(* CODESYS project Elevator_Control.project

Project tree, tasks and I/O mapping:
  Device : CODESYS Control Win V3, CODESYS, version 3.5.21.0
    application Application
      libraries: Standard, 3.5.18.0 (System)
      task MainTask (cyclic, interval 70 ms, priority 1) calls PLC_PRG, Simulation, GA_Collector
      task VISU_TASK (cyclic, interval 100 ms, priority 31) calls VisuElems.Visu_Prg
      global variables GVL
      visualisation Visualization
      program Simulation [ST]
      program GA_Collector [FBD]
      program PLC_PRG [SFC]: _aOpeningDoor_exit, _aCallsHMI_active, _aClosingDoor_active_1, _aClosingDoor_exit_1, _aOpeningDoor_active_1, _aOpenDoor_active, _aClosingDoor_exit_1_1_1_1_1, _aHoming_exit, _aHoming_active, _aOpeningDoor_active_1_1, _aOpeningDoor_exit_1, _aClosingDoor1_exit, _aClosingDoor1_active, _aClosingDoor_active_1_1_1_1_1, _aOpenDoor_exit, _aOpenDoor1_active, _aOpenDoor1_exit, _aTargetMoveStart_active, _aTargetMoveStart_exit, _aOpenDoor2_active, _aOpenDoor2_exit, _aResetCalls_active
      ENUMs/
        GAs/
          data type State_GA
          data type Action_State
          data type DoWhats_Closing
          data type DoWhats_Opening
          data type DoWhats_Motor
        data type Fault
        data type SensorSequence
      GAs/
        function block Opening_GA [SFC]: _aInit_active, _aReady_active, _aBusy_active, _aOpeningDoor_active, _aEnd_active, _aEnd_exit, _aOpeningDoor_exit
        function block Closing_GA [SFC]: _aInit_active, _aCheckPresence_active, _aBusy_active, _aClosingDoor_active, _aClosingDoor_exit, _aEnd_active, _aEnd_exit, _aReady_active_1
        function block Motor_GA [SFC]: _aBusy_active, _aEnd_Cycle_active, _aEnd_INIT_exit, _aInit_active, _aReady_active, _aEnd_Cycle_exit, _aMotor_ON_active, _aSetting_Down_active, _aMovingElevator_active, _aSetting_Init_active, _aSetting_Up_active, _aUpdateFloor_active_1, _aEnd_INIT_active, _aChangeDirection_exit, _aChangeDirection_active, _aMovingElevator_exit, _aSequenceCheck_active, _aMoveFast_entry_1, _aUpdateFloor_entry_1, _aInvertedSpeed1_active, _aInvertedSpeed_active_1, _aInvertedSpeed_exit, _aInvertedSpeed_entry
  text list GlobalTextList
*)

// Device/Application/ENUMs/GAs/State_GA
//{attribute 'qualified_only'}
//{attribute 'strict'}
TYPE State_GA :
(
	S_Init,
	S_Ready,
	S_Busy
);
END_TYPE

// Device/Application/ENUMs/GAs/Action_State
//{attribute 'qualified_only'}
//{attribute 'strict'}
TYPE Action_State :
(
	Do_Action,
	WaitDone,
	SetOpOk
);
END_TYPE

// Device/Application/ENUMs/Fault
//{attribute 'qualified_only'}
//{attribute 'strict'}
TYPE Fault :
(
	None,
	MagnetRamp,
	MagnetDeck
);
END_TYPE

// Device/Application/ENUMs/SensorSequence
//{attribute 'qualified_only'}
//{attribute 'strict'}
TYPE SensorSequence :
(
	Seq_Deck,
	Seq_Ramp1,
	Seq_Ramp2,
	Seq_Fault
);
END_TYPE

// Device/Application/ENUMs/GAs/DoWhats_Closing
//{attribute 'qualified_only'}
//{attribute 'strict'}
TYPE DoWhats_Closing :
(
	Do_CloseDoor
);
END_TYPE

// Device/Application/ENUMs/GAs/DoWhats_Opening
//{attribute 'qualified_only'}
//{attribute 'strict'}
TYPE DoWhats_Opening :
(
	Do_OpenDoor
);
END_TYPE

// Device/Application/ENUMs/GAs/DoWhats_Motor
//{attribute 'qualified_only'}
//{attribute 'strict'}
TYPE DoWhats_Motor :
(
	Do_Up,
	Do_Down, 
	Do_Inizialization
);
END_TYPE

// Device/Application/GVL
//{attribute 'qualified_only'}
VAR_GLOBAL
(* Elevator managing variables*)
	Open: BOOL;				(* Sensor: the door is fully open*)
	Closed: BOOL;			(* Sensor: the door is fully closed*)
	LimitDown: BOOL;		(* Sensor: lower limit sensor, if TRUE the lift has reached the lower limit*)
	LimitUp: BOOL;			(* Sensor: upper limit sensor, if TRUE the lift has reached the upper limit*)
	DeckSensor: BOOL;		(* Sensor: if TRUE the cab is in proximity of a deck*)
	RampSensor: BOOL;		(* Sensor: if TRUE the cab is in proximity of a ramp*)
	Presence :BOOL; 		(* Sensor: if TRUE something blocks the door photocell*)
	Emergency: BOOL;		(* Input: if TRUE the emergency button has been pressed*)

	Closing: BOOL;			(* Actuator: if TRUE the door starts closing*)
	Opening: BOOL;			(* Actuator: the door starts opening*)
	Motor_on: BOOL;			(* Actuator: if TRUE the lift pulley motor start moving*)
	Up: BOOL;				(* Actuator parameter: if TRUE the lift moves upward, downward otherwise*)
	Vel: BOOL;				(* Actuator parameter: motor speed, if TRUE high speed, low speed otherwise*)


	Current: INT;  			(* Visualization: variable used to storage the current deck*)
    Destination: INT;		(* Visualization: variable used to storage the the destination deck*)
	EmergencyVis: BOOL; 	(* Visualization: if TRUE the emergency light is turned on*)

	InitialDeck: INT := 1;	(* Only for simulation: variable used to define the initial deck*)
	InitCycle: BOOL := FALSE;(* Only for simulation: used to execute the instruction at the first cycle*)
	Height: INT;			(* Only for simulation: elevator height*)
	DeckRest: INT;        	(* Only for simulation: division rest for generating deck sensor*)
	Memory: INT;
	RampRest: INT;			(* Only for simulation: division rest for generating the ramp position*)
	MemoryR: INT;
	Door: INT;				(* Only for simulation: to visualize the closing of the door*)
	Displacement: INT;		(* Only for simulation: lift displacement, dependent on the motor speed*)

 (*Inputs: internal panel variables*)
	PG: BOOL;
	P1: BOOL;
	P2: BOOL;
	P3: BOOL;
	P4: BOOL;
	P5: BOOL;
	P6: BOOL;
	P7: BOOL;

(*Visualization: internal panel variables used to turn on the LED*)
	PGVis: BOOL;
	P1Vis: BOOL;
	P2Vis: BOOL;
	P3Vis: BOOL;
	P4Vis: BOOL;
	P5Vis: BOOL;
	P6Vis: BOOL;
	P7Vis: BOOL;

(*Inputs: external panel variables*)
	UpDeckG: BOOL;
	UpDeck1: BOOL;
	UpDeck2: BOOL;
	UpDeck3: BOOL;
	UpDeck4: BOOL;
	UpDeck5: BOOL;
	UpDeck6: BOOL;
	DownDeck7: BOOL;
	DownDeck6: BOOL;
	DownDeck5: BOOL;
	DownDeck4: BOOL;
	DownDeck3: BOOL;
	DownDeck2: BOOL;
	DownDeck1: BOOL;

(*Visualization: external panel variables used to turn on the LED*)
	UpDeckGVis: BOOL;
	UpDeck1Vis: BOOL;
	UpDeck2Vis: BOOL;
	UpDeck3Vis: BOOL;
	UpDeck4Vis: BOOL;
	UpDeck5Vis: BOOL;
	UpDeck6Vis: BOOL;
	DownDeck7Vis: BOOL;
	DownDeck6Vis: BOOL;
	DownDeck5Vis: BOOL;
	DownDeck4Vis: BOOL;
	DownDeck3Vis: BOOL;
	DownDeck2Vis: BOOL;
	DownDeck1Vis: BOOL;

(*Only for simulation: variables used to simulate the fault on deck sensor*)
	SensorG: BOOL;				(* if TRUE the magnetic information for deck G is lost and the deck sensor cannot become TRUE*)
	Sensor1: BOOL;				(* if TRUE the magnetic information for deck 1 is lost and the deck sensor cannot become TRUE*)
	Sensor2: BOOL;
	Sensor3: BOOL;
	Sensor4: BOOL;
	Sensor5: BOOL;
	Sensor6: BOOL;
	Sensor7: BOOL;
	FaultSensorAlarm: BOOL; 	(* Visulaization: if TRUE alerts the user of a deck sensor fault*)

(*Only for simulation: variables used to simulate the fault on ramp sensor*)
	RampGUp: BOOL;
	Ramp1Down: BOOL;
	Ramp1Up:BOOL;
	Ramp2Down: BOOL;
	Ramp2Up:BOOL;
	Ramp3Down: BOOL;
	Ramp3Up:BOOL;
	Ramp4Down: BOOL;
	Ramp4Up:BOOL;
	Ramp5Down: BOOL;
	Ramp5Up:BOOL;
	Ramp6Down: BOOL;
	Ramp6Up:BOOL;
	Ramp7Down: BOOL;
	FaultRampAlarm: BOOL; 		(* Visulaization: if TRUE alerts the user of a ramp sensor fault*)
	SensorGOK: BOOL;
	Sensor1OK: BOOL;
	Sensor2OK: BOOL;
	Sensor6OK: BOOL;
	Sensor3OK: BOOL;
	Sensor4OK: BOOL;
	Sensor5OK: BOOL;
	Sensor7OK: BOOL;
	RampGUpOK: BOOL;
	Ramp1DownOK: BOOL;
	Ramp1UpOK: BOOL;
	Ramp2DownOK: BOOL;
	Ramp2UpOK: BOOL;
	Ramp3DownOK: BOOL;
	Ramp3UpOK: BOOL;
	Ramp4DownOK: BOOL;
	Ramp4UpOK: BOOL;
	Ramp5DownOK: BOOL;
	Ramp5UpOK: BOOL;
	Ramp6DownOK: BOOL;
	Ramp6UpOK: BOOL;
	Ramp7DownOK: BOOL;
	Ramp7UpOK: BOOL;
	
	Closing_GA_0: Closing_GA;
	Opening_GA_0: Opening_GA;
	Motor_GA_0: Motor_GA;
END_VAR

// Device/Application/PLC_PRG
PROGRAM PLC_PRG
VAR
	A_State: Action_State := Do_Action;
	OpOk: BOOL;
	IntPanel : ARRAY [0..7] OF BOOL;
	ExtPanelUP : ARRAY [0..6] OF BOOL;
	ExtPanelDOWN : ARRAY [1..7] OF BOOL;
	CallInt : ARRAY[0..7] OF BOOL; //chiamate interne
	CallUp : ARRAY[0..6] OF BOOL;     //chiamate esterne vs alto
	CallDown : ARRAY[1..7] OF BOOL;   //chiamate esterne vs basso   
	i : INT;
END_VAR

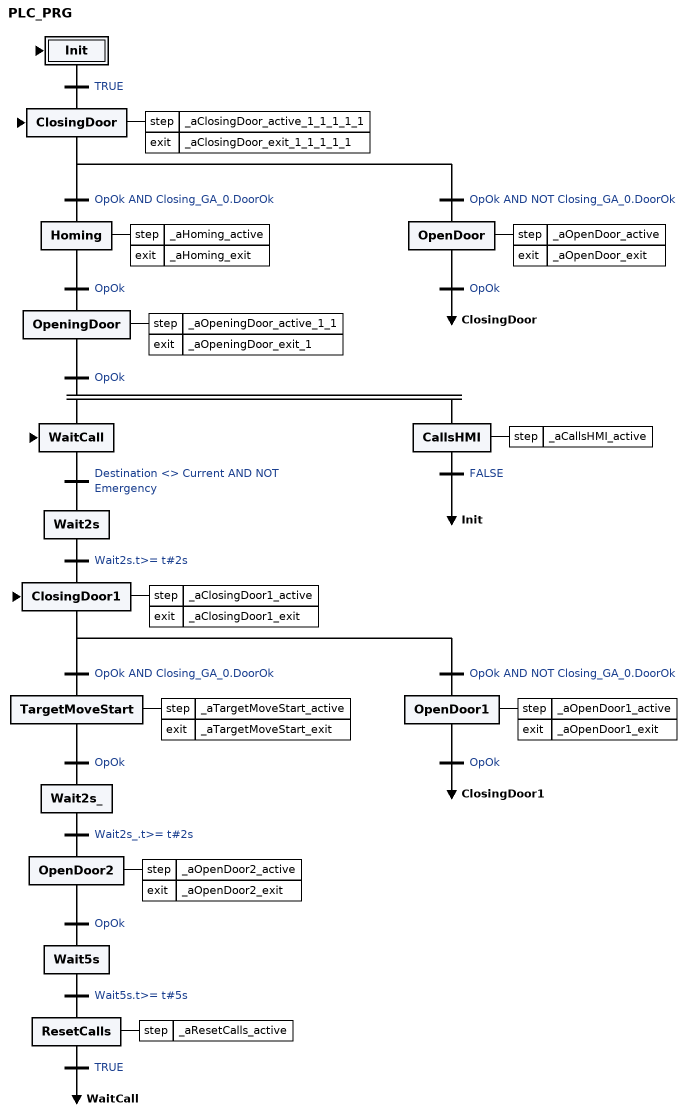
INITIAL_STEP Init:
END_STEP
TRANSITION FROM Init TO ClosingDoor
    := TRUE;
END_TRANSITION
STEP ClosingDoor:
    _aClosingDoor_active_1_1_1_1_1(N);  // step action
    _aClosingDoor_exit_1_1_1_1_1(P0);  // exit action
END_STEP
TRANSITION FROM ClosingDoor TO Homing
    := OpOk AND Closing_GA_0.DoorOk;
END_TRANSITION
TRANSITION FROM ClosingDoor TO OpenDoor
    := OpOk AND NOT Closing_GA_0.DoorOk;
END_TRANSITION
STEP OpenDoor:
    _aOpenDoor_active(N);  // step action
    _aOpenDoor_exit(P0);  // exit action
END_STEP
TRANSITION FROM OpenDoor TO ClosingDoor
    := OpOk;
END_TRANSITION
STEP Homing:
    _aHoming_active(N);  // step action
    _aHoming_exit(P0);  // exit action
END_STEP
TRANSITION FROM Homing TO OpeningDoor
    := OpOk;
END_TRANSITION
STEP OpeningDoor:
    _aOpeningDoor_active_1_1(N);  // step action
    _aOpeningDoor_exit_1(P0);  // exit action
END_STEP
TRANSITION FROM OpeningDoor TO (WaitCall, CallsHMI)
    := OpOk;
END_TRANSITION
STEP WaitCall:
END_STEP
STEP CallsHMI:
    _aCallsHMI_active(N);  // step action
END_STEP
TRANSITION FROM CallsHMI TO Init
    := FALSE;
END_TRANSITION
TRANSITION FROM WaitCall TO Wait2s
    := Destination <> Current AND NOT Emergency;
END_TRANSITION
STEP Wait2s:
END_STEP
TRANSITION FROM Wait2s TO ClosingDoor1
    := Wait2s.t>= t#2s;
END_TRANSITION
STEP ClosingDoor1:
    _aClosingDoor1_active(N);  // step action
    _aClosingDoor1_exit(P0);  // exit action
END_STEP
TRANSITION FROM ClosingDoor1 TO TargetMoveStart
    := OpOk AND Closing_GA_0.DoorOk;
END_TRANSITION
TRANSITION FROM ClosingDoor1 TO OpenDoor1
    := OpOk AND NOT Closing_GA_0.DoorOk;
END_TRANSITION
STEP OpenDoor1:
    _aOpenDoor1_active(N);  // step action
    _aOpenDoor1_exit(P0);  // exit action
END_STEP
TRANSITION FROM OpenDoor1 TO ClosingDoor1
    := OpOk;
END_TRANSITION
STEP TargetMoveStart:
    _aTargetMoveStart_active(N);  // step action
    _aTargetMoveStart_exit(P0);  // exit action
END_STEP
TRANSITION FROM TargetMoveStart TO Wait2s_
    := OpOk;
END_TRANSITION
STEP Wait2s_:
END_STEP
TRANSITION FROM Wait2s_ TO OpenDoor2
    := Wait2s_.t>= t#2s;
END_TRANSITION
STEP OpenDoor2:
    _aOpenDoor2_active(N);  // step action
    _aOpenDoor2_exit(P0);  // exit action
END_STEP
TRANSITION FROM OpenDoor2 TO Wait5s
    := OpOk;
END_TRANSITION
STEP Wait5s:
END_STEP
TRANSITION FROM Wait5s TO ResetCalls
    := Wait5s.t>= t#5s;
END_TRANSITION
STEP ResetCalls:
    _aResetCalls_active(N);  // step action
END_STEP
TRANSITION FROM ResetCalls TO WaitCall
    := TRUE;
END_TRANSITION

ACTION _aOpeningDoor_exit:
OpOk := FALSE;
A_State := Do_Action;
END_ACTION

ACTION _aCallsHMI_active:
// Mappatura dei tasti della pulsantiera interna sui piani
IntPanel[0] := PG;
IntPanel[1] := P1;
IntPanel[2] := P2;
IntPanel[3] := P3;
IntPanel[4] := P4;
IntPanel[5] := P5;
IntPanel[6] := P6;
IntPanel[7] := P7;

//Gestione delle richieste interne
FOR i := 0 TO 7 DO
	IF IntPanel[i] THEN
		CallInt[i] := TRUE;   	//Salva richiesta interna attiva
	END_IF
	IF (Current = i) AND Open THEN
		CallInt[i] := FALSE;   // Cancella richiesta se cabina è ferma al piano e porte aperte
	END_IF
END_FOR

// Mappatura dei tasti di salita della pulsantiera esterna
ExtPanelUP[0] := UpDeckG;
ExtPanelUP[1] := UpDeck1;
ExtPanelUP[2] := UpDeck2;
ExtPanelUP[3] := UpDeck3;
ExtPanelUP[4] := UpDeck4;
ExtPanelUP[5] := UpDeck5;
ExtPanelUP[6] := UpDeck6;

//Gestione delle richieste esterne verso l'alto
FOR i:= 0 TO 6 DO
	IF ExtPanelUP[i] THEN 
		CallUp[i] := TRUE;        
	END_IF;
	IF (Current = i) AND Open THEN
	CallUp[i] := FALSE;           
	END_IF
END_FOR

// Mappatura dei tasti di discesa della pulsantiera esterna
ExtPanelDOWN[1] := DownDeck1;
ExtPanelDOWN[2] := DownDeck2;
ExtPanelDOWN[3] := DownDeck3;
ExtPanelDOWN[4] := DownDeck4;
ExtPanelDOWN[5] := DownDeck5;
ExtPanelDOWN[6] := DownDeck6;
ExtPanelDOWN[7] := DownDeck7;

// Gestione delle richieste esterne verso il basso
FOR i := 1 TO 7 DO
	IF ExtPanelDown[i] THEN
		CallDown[i] := TRUE;
	END_IF
	IF (Current = i) AND Open THEN
	CallDown[i] := FALSE;
	END_IF
END_FOR

//Aggiornamento LED interni in base alle richieste
PGVis := CallInt[0];
P1Vis := CallInt[1];
P2Vis := CallInt[2];
P3Vis := CallInt[3];
P4Vis := CallInt[4];
P5Vis := CallInt[5];
P6Vis := CallInt[6];
P7Vis := CallInt[7];

//Aggiornamento LED esterni salita
UpDeckGVis := CallUp[0];
UpDeck1Vis := CallUp[1];
UpDeck2Vis := CallUp[2];
UpDeck3Vis := CallUp[3];
UpDeck4Vis := CallUp[4];
UpDeck5Vis := CallUp[5];
UpDeck6Vis := CallUp[6];

//Aggiornamento LED esterni discesa
DownDeck1Vis := CallDown[1];
DownDeck2Vis := CallDown[2];
DownDeck3Vis := CallDown[3];
DownDeck4Vis := CallDown[4];
DownDeck5Vis := CallDown[5];
DownDeck6Vis := CallDown[6];
DownDeck7Vis := CallDown[7]; 

// Gestione indicatori emergency e faults
IF Emergency THEN
	EmergencyVis := TRUE;
ELSE
	EmergencyVis := FALSE;
END_IF

IF Motor_GA_0.Fault_State = MagnetDeck THEN
	FaultSensorAlarm := TRUE;
ELSE
	FaultSensorAlarm := FALSE;
END_IF

IF Motor_GA_0.Fault_State = MagnetRamp THEN
	FaultRampAlarm := TRUE;
ELSE
	FaultRampAlarm := FALSE;
END_IF

//Scansione verso l’alto per trovare una destinazione valida
FOR i := Current+1 TO 7 DO        
    IF (CallInt[i] OR CallUp[i]) AND NOT Emergency THEN
		IF Motor_GA_0.Fault_State = None THEN
        	Destination := i;
		ELSIF (Motor_GA_0.Fault_State = MagnetRamp) OR (Motor_GA_0.Fault_State = MagnetDeck) THEN         
			Destination := Current;
		END_IF
	ELSIF (CallInt[i] OR CallUp[i]) AND Emergency THEN
		Destination := Current;
        RETURN;
    END_IF;
END_FOR;

IF Current <> -1 THEN                            //Il current va a -1 per un certo istante quando vi è un fault sul piano G
FOR i := Current+1 TO 7 DO                       //CallDown va da 1 a 7 => per current = -1 si avrebbe i = 0 dando così errore
    IF (CallDown[i]) AND NOT Emergency THEN      //Codice come quello sopra che consente scansione verso l'alto anche per chiamate con freccia in basso
		IF Motor_GA_0.Fault_State = None THEN
        	Destination := i;
		ELSIF (Motor_GA_0.Fault_State = MagnetRamp) OR (Motor_GA_0.Fault_State = MagnetDeck) THEN         
			Destination := Current;
		END_IF
	ELSIF (CallInt[i] OR CallUp[i]) AND Emergency THEN
		Destination := Current;
        RETURN;
    END_IF;
END_FOR;
END_IF

// Se non ci sono richieste in alto, cerca verso il basso
FOR i :=  Current-1 TO 1 BY -1 DO      
    IF (CallInt[i] OR CallDown[i] OR CallUp[i]) AND NOT Emergency THEN
		IF Motor_GA_0.Fault_State = None THEN
	        Destination := i;
		ELSIF (Motor_GA_0.Fault_State = MagnetRamp) OR (Motor_GA_0.Fault_State = MagnetDeck) THEN         
			Destination := Current;
			END_IF;
	ELSIF (CallInt[i] OR CallDown[i]) AND Emergency THEN
		Destination := Current;
        RETURN;
    END_IF;
END_FOR;  

// Controllo separato per piano 0. Non è presente CallDown[0], quindi non può essere incluso nel ciclo generale.
// In tal modo il ciclo for precedente non va in errore.

 IF (CallInt[0] OR CallUp[0]) AND NOT Emergency THEN
	IF Motor_GA_0.Fault_State = None THEN
	        Destination := 0;
	ELSIF (Motor_GA_0.Fault_State = MagnetRamp) OR (Motor_GA_0.Fault_State = MagnetDeck) THEN        
			Destination := Current;
 	END_IF;
ELSIF (CallInt[0] OR CallUp[0]) AND Emergency THEN
	Destination := Current;
    RETURN;
END_IF;
END_ACTION

ACTION _aClosingDoor_active_1:
CASE A_State OF
	Do_Action: IF Closing_GA_0.State = S_Ready THEN
		Closing_GA_0.Do_ := TRUE;
		Closing_GA_0.DoWhat := Do_CloseDoor;
		A_State := WaitDone;
	END_IF
	WaitDone: IF Closing_GA_0.Done AND Closing_GA_0.State = S_Busy THEN
			  	Closing_GA_0.Do_ := FALSE;
				A_State := SetOpOk;
				END_IF	
	SetOpOk:  IF NOT Closing_GA_0.Done THEN 
		      OpOk:= TRUE;
		      END_IF
END_CASE
END_ACTION

ACTION _aClosingDoor_exit_1:
OpOk := FALSE;
A_State := Do_Action;
END_ACTION

ACTION _aOpeningDoor_active_1:
CASE A_State OF
	Do_Action: IF Opening_GA_0.State = S_Ready THEN
		Opening_GA_0.Do_ := TRUE;
		Opening_GA_0.DoWhat := Do_OpenDoor;
		A_State := WaitDone;
	END_IF
	WaitDone: IF Opening_GA_0.Done AND Opening_GA_0.State = S_Busy THEN
			  	Opening_GA_0.Do_ := FALSE;
				A_State := SetOpOk;
				END_IF	
	SetOpOk:  IF NOT Opening_GA_0.Done THEN 
		      OpOk:= TRUE;
		      END_IF
END_CASE
END_ACTION

ACTION _aOpenDoor_active:
CASE A_State OF
	Do_Action: IF Opening_GA_0.State = S_Ready THEN
		Opening_GA_0.Do_ := TRUE;
		Opening_GA_0.DoWhat := Do_OpenDoor;
		A_State := WaitDone;
	END_IF
	WaitDone: IF Opening_GA_0.Done AND Opening_GA_0.State = S_Busy THEN
			  	Opening_GA_0.Do_ := FALSE;
				A_State := SetOpOk;
				END_IF	
	SetOpOk:  IF NOT Opening_GA_0.Done THEN 
		      OpOk:= TRUE;
		      END_IF
END_CASE
END_ACTION

ACTION _aClosingDoor_exit_1_1_1_1_1:
OpOk := FALSE;
A_State := Do_Action;
END_ACTION

ACTION _aHoming_exit:
OpOk := FALSE;
A_State := Do_Action;
END_ACTION

ACTION _aHoming_active:
CASE A_State OF
	Do_Action: IF Motor_GA_0.State = S_Ready THEN
		Motor_GA_0.Do_ := TRUE;
		Motor_GA_0.DoWhat := Do_Inizialization;
		A_State := WaitDone;
	END_IF
	WaitDone: IF Motor_GA_0.Done AND Motor_GA_0.State = S_Busy THEN
			  	Motor_GA_0.Do_ := FALSE;
				A_State := SetOpOk;
				END_IF	
	SetOpOk:  IF NOT Motor_GA_0.Done THEN 
		      OpOk:= TRUE;
		      END_IF
END_CASE
END_ACTION

ACTION _aOpeningDoor_active_1_1:
CASE A_State OF
	Do_Action: IF Opening_GA_0.State = S_Ready THEN
		Opening_GA_0.Do_ := TRUE;
		Opening_GA_0.DoWhat := Do_OpenDoor;
		A_State := WaitDone;
	END_IF
	WaitDone: IF Opening_GA_0.Done AND Opening_GA_0.State = S_Busy THEN
			  	Opening_GA_0.Do_ := FALSE;
				A_State := SetOpOk;
				END_IF	
	SetOpOk:  IF NOT Opening_GA_0.Done THEN 
		      OpOk:= TRUE;
		      END_IF
END_CASE
END_ACTION

ACTION _aOpeningDoor_exit_1:
OpOk := FALSE;
A_State := Do_Action;
END_ACTION

ACTION _aClosingDoor1_exit:
OpOk := FALSE;
A_State := Do_Action;
END_ACTION

ACTION _aClosingDoor1_active:
CASE A_State OF
	Do_Action: IF Closing_GA_0.State = S_Ready THEN
		Closing_GA_0.Do_ := TRUE;
		Closing_GA_0.DoWhat := Do_CloseDoor;
		A_State := WaitDone;
	END_IF
	WaitDone: IF Closing_GA_0.Done AND Closing_GA_0.State = S_Busy THEN
			  	Closing_GA_0.Do_ := FALSE;
				A_State := SetOpOk;
				END_IF	
	SetOpOk:  IF NOT Closing_GA_0.Done THEN 
		      OpOk:= TRUE;
		      END_IF
END_CASE
END_ACTION

ACTION _aClosingDoor_active_1_1_1_1_1:
CASE A_State OF
	Do_Action: IF Closing_GA_0.State = S_Ready THEN
		Closing_GA_0.Do_ := TRUE;
		Closing_GA_0.DoWhat := Do_CloseDoor;
		A_State := WaitDone;
	END_IF
	WaitDone: IF Closing_GA_0.Done AND Closing_GA_0.State = S_Busy THEN
			  	Closing_GA_0.Do_ := FALSE;
				A_State := SetOpOk;
				END_IF	
	SetOpOk:  IF NOT Closing_GA_0.Done THEN 
		      OpOk:= TRUE;
		      END_IF
END_CASE
END_ACTION

ACTION _aOpenDoor_exit:
OpOk := FALSE;
A_State := Do_Action;
END_ACTION

ACTION _aOpenDoor1_active:
CASE A_State OF
	Do_Action: IF Opening_GA_0.State = S_Ready THEN
		Opening_GA_0.Do_ := TRUE;
		Opening_GA_0.DoWhat := Do_OpenDoor;
		A_State := WaitDone;
	END_IF
	WaitDone: IF Opening_GA_0.Done AND Opening_GA_0.State = S_Busy THEN
			  	Opening_GA_0.Do_ := FALSE;
				A_State := SetOpOk;
				END_IF	
	SetOpOk:  IF NOT Opening_GA_0.Done THEN 
		      OpOk:= TRUE;
		      END_IF
END_CASE
END_ACTION

ACTION _aOpenDoor1_exit:
OpOk := FALSE;
A_State := Do_Action;
END_ACTION

ACTION _aTargetMoveStart_active:
CASE A_State OF
	Do_Action:
		 IF Motor_GA_0.State = S_Ready THEN    						
		   IF Destination > Current THEN 	// Determina la direzione
		Motor_GA_0.DoWhat := Do_Up;			
		ELSIF Destination < Current THEN
		Motor_GA_0.DoWhat := Do_Down;
		END_IF
		Motor_GA_0.Do_ := TRUE;	
		A_State := WaitDone;          	   
			
		END_IF
	WaitDone: 
		// Controllo delle chiamate "al volo" durante il tragitto
			// se sto salendo
			IF Motor_GA_0.DoWhat = Do_Up  THEN    
				FOR i := Current+1 TO Destination-1 DO    		// Cerca eventuale nuova chiamata interna/esterna verso l'alto più vicina
					IF CallInt[i] OR CallUp[i] OR CallDown[i] THEN
						Destination := i;             	 	    // Cambio destinazione se trovo una chiamata più urgente
						EXIT;                             
					END_IF;
				END_FOR;
			
			// se sto scendendo
			ELSIF Motor_GA_0.DoWhat = Do_Down  THEN
				FOR i := Current-1 TO Destination+1 BY -1 DO     // Cerca eventuale nuova chiamata interna/esterna verso il basso più vicina
					IF CallInt[i] OR CallDown[i] OR CallUp[i] THEN
						Destination := i;                        // Cambio destinazione se trovo una chiamata più urgente
						EXIT;
					END_IF;
				END_FOR;
			END_IF;

			IF Motor_GA_0.Done AND Motor_GA_0.State = S_Busy THEN
			  Motor_GA_0.Do_ := FALSE;
				A_State := SetOpOk;
				END_IF	
	SetOpOk:  IF NOT Motor_GA_0.Done THEN 
		      OpOk:= TRUE;
		      END_IF
END_CASE
END_ACTION

ACTION _aTargetMoveStart_exit:
OpOk := FALSE;
A_State := Do_Action;
END_ACTION

ACTION _aOpenDoor2_active:
CASE A_State OF
	Do_Action: IF Opening_GA_0.State = S_Ready THEN
		Opening_GA_0.Do_ := TRUE;
		Opening_GA_0.DoWhat := Do_OpenDoor;
		A_State := WaitDone;
	END_IF
	WaitDone: IF Opening_GA_0.Done AND Opening_GA_0.State = S_Busy THEN
			  	Opening_GA_0.Do_ := FALSE;
				A_State := SetOpOk;
				END_IF	
	SetOpOk:  IF NOT Opening_GA_0.Done THEN 
		      OpOk:= TRUE;
		      END_IF
END_CASE
END_ACTION

ACTION _aOpenDoor2_exit:
OpOk := FALSE;
A_State := Do_Action;
END_ACTION

ACTION _aResetCalls_active:
IF Open THEN
    
    CallInt[Current] := FALSE;		  // Reset della chiamata interna al piano attuale, sempre valido
   
    IF Current < 7 THEN
        CallUp[Current] := FALSE;     // Reset della chiamata esterna in salita (solo se non siamo all’ultimo piano)
    END_IF;

    IF Current > 0 THEN
        CallDown[Current] := FALSE;   // Reset della chiamata esterna in discesa (solo se non siamo al piano 0)
    END_IF;
END_IF;
END_ACTION

END_PROGRAM

// Device/Application/Simulation
PROGRAM Simulation
VAR
END_VAR

(* Initial position of the cab inside the hoistway. It is executed only at the first cycle.  *)
IF NOT GVL.InitCycle THEN
			GVL.InitCycle := TRUE ;
			GVL.Height := 20 * GVL.InitialDeck;
		    GVL.Door := 0;
			GVL.Current := GVL.Height / 20;
END_IF;

(* Elevator management, these instructions are executed each cycle time*)

(* Elevator door control. *)
IF GVL.Closing THEN
	GVL.Door := GVL.Door + 1;		(*Closing door management*)
	GVL.Open := FALSE;
END_IF

IF GVL.Door >= 60 THEN						(* Closed door limit*)
	GVL.Closed := TRUE;
END_IF

IF GVL.Opening THEN
	GVL.Door := GVL.Door - 1; 	(* Opening door management*)
	GVL.Closed := FALSE;
END_IF

IF GVL.Door <= 0 THEN							(* Open door limit*)
	GVL.Open := TRUE;
END_IF


(* Maximum and minimum management in the door simulation*)
IF GVL.Door < 0 THEN
	 GVL.Door := 0;
END_IF

IF GVL.Door > 60 THEN
	GVL.Door := 60;
END_IF


(* Control of the cab position inside the hostway. *)
(* Displacement definition for graphic visualization*)
IF GVL.Vel THEN 
	GVL.Displacement := 2;
ELSE 
	GVL.Displacement := 1;
END_IF


(* Height modification relying on direction and speed*)
IF GVL.Motor_on AND GVL.Up THEN
	GVL.Height := GVL.Height + GVL.Displacement;
	GVL.LimitDown := FALSE;
END_IF

IF GVL.Motor_on AND NOT GVL.Up THEN
	GVL.Height := GVL.Height - GVL.Displacement;
	GVL.LimitUp := FALSE;
END_IF


(* Limits for visualization*)
IF GVL.Height < -20 THEN
	GVL.Height := -20;
END_IF

IF GVL.Height > 160 THEN
	GVL.Height := 160;
END_IF

(* Limit sensors management*)
IF GVL.Height <= -10 THEN
	GVL.LimitDown := TRUE;
END_IF

IF GVL.Height >= 150 THEN
	 GVL.LimitUp := TRUE;
END_IF


(*-------------------------------------------------------------------*)
(*  Fault Management (Deck and Ramp Sensors)   *)
(*-------------------------------------------------------------------*)
(* Deck Sensor*)
(* Range of value where the deck sensor is active*)
IF ((GVL.Height >= -1) AND (GVL.Height <= 1)) THEN
	GVL.SensorGOK := TRUE;
ELSE  
	GVL.SensorGOK := FALSE;
END_IF

IF ((GVL.Height >= 20-1) AND (GVL.Height <= 20+1)) THEN
	GVL.Sensor1OK := TRUE;
ELSE  
	GVL.Sensor1OK := FALSE;
END_IF

IF ((GVL.Height >= 40-1) AND (GVL.Height <= 40+1)) THEN
	GVL.Sensor2OK := TRUE;
ELSE  
	GVL.Sensor2OK := FALSE;
END_IF

IF ((GVL.Height >= 60-1) AND (GVL.Height <= 60+1)) THEN
	GVL.Sensor3OK := TRUE;
ELSE  
	GVL.Sensor3OK := FALSE;
END_IF

IF ((GVL.Height >= 80-1) AND (GVL.Height <= 80+1)) THEN
	GVL.Sensor4OK := TRUE;
ELSE  
	GVL.Sensor4OK := FALSE;
END_IF

IF ((GVL.Height >= 100-1) AND (GVL.Height <= 100+1)) THEN
	GVL.Sensor5OK := TRUE;
ELSE   
	GVL.Sensor5OK := FALSE;
END_IF

IF ((GVL.Height >= 120-1) AND (GVL.Height <= 120+1)) THEN
	GVL.Sensor6OK := TRUE;
ELSE  
	GVL.Sensor6OK := FALSE;
END_IF

IF ((GVL.Height >= 140-1) AND (GVL.Height <= 140+1)) THEN
	GVL.Sensor7OK := TRUE;
ELSE  
	GVL.Sensor7OK := FALSE;
END_IF

GVL.DeckSensor := (GVL.SensorGOK AND NOT GVL.SensorG) OR
				    (GVL.Sensor1OK AND NOT GVL.Sensor1) OR
				    (GVL.Sensor2OK AND NOT GVL.Sensor2) OR
				    (GVL.Sensor3OK AND NOT GVL.Sensor3) OR
				    (GVL.Sensor4OK AND NOT GVL.Sensor4) OR
				    (GVL.Sensor5OK AND NOT GVL.Sensor5) OR
				    (GVL.Sensor6OK AND NOT GVL.Sensor6) OR
				    (GVL.Sensor7OK AND NOT GVL.Sensor7);

(* Ramp Sensor*)
(* Range of value where the ramp sensor is active*)
IF ((GVL.Height >= 5-1) AND (GVL.Height <= 5+1)) THEN
	GVL.RampGUpOK := TRUE;
ELSE 
	GVL.RampGUpOK := FALSE;
END_IF

(* Ramp close to deck 1*)
IF ((GVL.Height >= 15-1) AND (GVL.Height <= 15+1)) THEN
	GVL.Ramp1DownOK := TRUE;
ELSE 
	GVL.Ramp1DownOK := FALSE;
END_IF

IF ((GVL.Height >= 25-1) AND (GVL.Height <= 25+1)) THEN
	GVL.Ramp1UpOK := TRUE;
ELSE 
	GVL.Ramp1UpOK := FALSE;
END_IF

(* Ramp close to deck 2*)
IF ((GVL.Height >= 35-1) AND (GVL.Height <= 35+1)) THEN
	GVL.Ramp2DownOK := TRUE;
ELSE 
	GVL.Ramp2DownOK := FALSE;
END_IF

IF ((GVL.Height >= 45-1) AND (GVL.Height <= 45+1)) THEN
	GVL.Ramp2UpOK := TRUE;
ELSE 
	GVL.Ramp2UpOK := FALSE;
END_IF

(*Ramp close to deck  3*)
IF ((GVL.Height >= 55-1) AND (GVL.Height <= 55+1)) THEN
	GVL.Ramp3DownOK := TRUE;
ELSE 
	GVL.Ramp3DownOK := FALSE;
END_IF

IF ((GVL.Height >= 65-1) AND (GVL.Height <= 65+1)) THEN
	GVL.Ramp3UpOK := TRUE;
ELSE 
	GVL.Ramp3UpOK := FALSE;
END_IF

(* Ramp close to deck  4*)
IF ((GVL.Height >= 75-1) AND (GVL.Height <= 75+1)) THEN
	GVL.Ramp4DownOK := TRUE;
ELSE 
	GVL.Ramp4DownOK := FALSE;
END_IF

IF ((GVL.Height >= 85-1) AND (GVL.Height <= 85+1)) THEN
	GVL.Ramp4UpOK := TRUE;
ELSE 
	GVL.Ramp4UpOK:=FALSE;
END_IF

(* Ramp close to deck  5*)
IF ((GVL.Height >= 95-1) AND (GVL.Height <= 95+1)) THEN
	GVL.Ramp5DownOK := TRUE;
ELSE 
	GVL.Ramp5DownOK := FALSE;
END_IF

IF ((GVL.Height >= 105-1) AND (GVL.Height <= 105+1)) THEN
	GVL.Ramp5UpOK := TRUE;
ELSE
	GVL.Ramp5UpOK := FALSE;
END_IF

(* Ramp close to deck  6*)
IF ((GVL.Height >= 115-1) AND (GVL.Height <= 115+1)) THEN
	GVL.Ramp6DownOK := TRUE;
ELSE 
	GVL.Ramp6DownOK := FALSE;
END_IF

IF ((GVL.Height >= 125-1) AND (GVL.Height <= 125+1)) THEN
	GVL.Ramp6UpOK := TRUE;
ELSE 
	GVL.Ramp6UpOK := FALSE;
END_IF

(* Ramp close to deck  7*)
IF ((GVL.Height >= 135-1) AND (GVL.Height <= 135+1)) THEN
	GVL.Ramp7DownOK := TRUE;
ELSE 
	GVL.Ramp7DownOK := FALSE;
END_IF

GVL.RampSensor:=(GVL.RampGUpOK AND NOT GVL.RampGUp) OR 
								(GVL.Ramp1DownOK AND NOT GVL.Ramp1Down ) OR 
								(GVL.Ramp1UpOK AND NOT GVL.Ramp1Up ) OR
								(GVL.Ramp2DownOK AND NOT GVL.Ramp2Down ) OR 
								(GVL.Ramp2UpOK AND NOT GVL.Ramp2Up ) OR
								(GVL.Ramp3DownOK AND NOT GVL.Ramp3Down ) OR
 								(GVL.Ramp3UpOK AND NOT GVL.Ramp3Up ) OR
								(GVL.Ramp4DownOK AND NOT GVL.Ramp4Down ) OR
 								(GVL.Ramp4UpOK AND NOT GVL.Ramp4Up ) OR
								(GVL.Ramp5DownOK AND NOT GVL.Ramp5Down ) OR
 								(GVL.Ramp5UpOK AND NOT GVL.Ramp5Up ) OR
								(GVL.Ramp6DownOK AND NOT GVL.Ramp6Down ) OR
								(GVL.Ramp6UpOK AND NOT GVL.Ramp6Up ) OR
								(GVL.Ramp7DownOK AND NOT GVL.Ramp7Down );

END_PROGRAM

// Device/Application/GA_Collector
PROGRAM GA_Collector
VAR
END_VAR

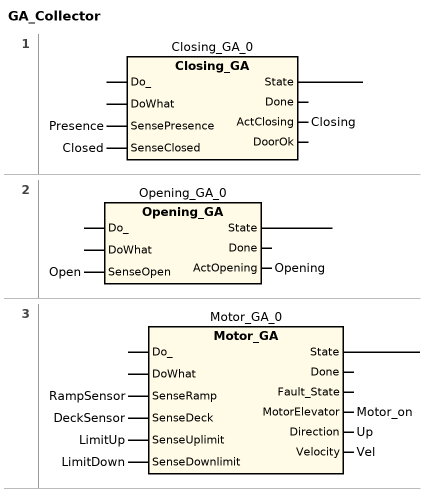
// NETWORK 1
Closing_GA_0(SensePresence := Presence, SenseClosed := Closed, ActClosing => Closing); // Closing_GA

// NETWORK 2
Opening_GA_0(SenseOpen := Open, ActOpening => Opening); // Opening_GA

// NETWORK 3
Motor_GA_0(
    SenseRamp := RampSensor,
    SenseDeck := DeckSensor,
    SenseUplimit := LimitUp,
    SenseDownlimit := LimitDown,
    MotorElevator => Motor_on,
    Direction => Up,
    Velocity => Vel); // Motor_GA

END_PROGRAM

// Device/Application/GAs/Closing_GA
FUNCTION_BLOCK Closing_GA
VAR_INPUT
	Do_: BOOL;
	DoWhat: DoWhats_Closing;
	SensePresence: BOOL;
	SenseClosed: BOOL;
END_VAR
VAR_OUTPUT
	State: State_GA;
	Done: BOOL;
	ActClosing: BOOL;
	DoorOk: BOOL;
END_VAR
VAR
END_VAR

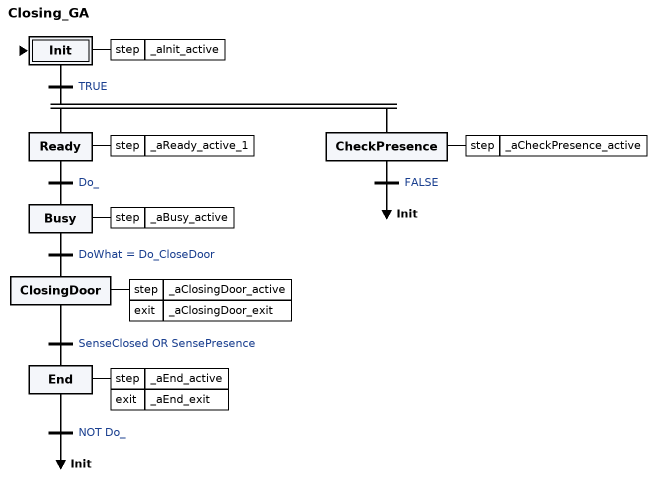
INITIAL_STEP Init:
    _aInit_active(N);  // step action
END_STEP
TRANSITION FROM Init TO (Ready, CheckPresence)
    := TRUE;
END_TRANSITION
STEP Ready:
    _aReady_active_1(N);  // step action
END_STEP
STEP CheckPresence:
    _aCheckPresence_active(N);  // step action
END_STEP
TRANSITION FROM CheckPresence TO Init
    := FALSE;
END_TRANSITION
TRANSITION FROM Ready TO Busy
    := Do_;
END_TRANSITION
STEP Busy:
    _aBusy_active(N);  // step action
END_STEP
TRANSITION FROM Busy TO ClosingDoor
    := DoWhat = Do_CloseDoor;
END_TRANSITION
STEP ClosingDoor:
    _aClosingDoor_active(N);  // step action
    _aClosingDoor_exit(P0);  // exit action
END_STEP
TRANSITION FROM ClosingDoor TO End
    := SenseClosed OR SensePresence;
END_TRANSITION
STEP End:
    _aEnd_active(N);  // step action
    _aEnd_exit(P0);  // exit action
END_STEP
TRANSITION FROM End TO Init
    := NOT Do_;
END_TRANSITION

ACTION _aInit_active:
State := S_Init;
END_ACTION

ACTION _aCheckPresence_active:
// controllo presenza passeggero 
// Se si ha DoorOk a FALSE, la politica blocca la chiusura porte.

IF NOT SensePresence THEN
	DoorOk := TRUE;
ELSE
	DoorOk := FALSE;
END_IF
END_ACTION

ACTION _aBusy_active:
State := S_Busy;
END_ACTION

ACTION _aClosingDoor_active:
ActClosing := TRUE;
END_ACTION

ACTION _aClosingDoor_exit:
ActClosing := FALSE;
END_ACTION

ACTION _aEnd_active:
Done := TRUE;
END_ACTION

ACTION _aEnd_exit:
Done := FALSE;
END_ACTION

ACTION _aReady_active_1:
State := S_Ready;
END_ACTION

END_FUNCTION_BLOCK

// Device/Application/GAs/Opening_GA
FUNCTION_BLOCK Opening_GA
VAR_INPUT
	Do_: BOOL;
	DoWhat: DoWhats_Opening;
	SenseOpen: BOOL;
END_VAR
VAR_OUTPUT
	State: State_GA;
	Done: BOOL;
	ActOpening: BOOL;
END_VAR
VAR
END_VAR

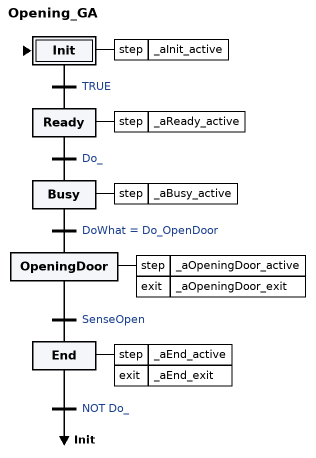
INITIAL_STEP Init:
    _aInit_active(N);  // step action
END_STEP
TRANSITION FROM Init TO Ready
    := TRUE;
END_TRANSITION
STEP Ready:
    _aReady_active(N);  // step action
END_STEP
TRANSITION FROM Ready TO Busy
    := Do_;
END_TRANSITION
STEP Busy:
    _aBusy_active(N);  // step action
END_STEP
TRANSITION FROM Busy TO OpeningDoor
    := DoWhat = Do_OpenDoor;
END_TRANSITION
STEP OpeningDoor:
    _aOpeningDoor_active(N);  // step action
    _aOpeningDoor_exit(P0);  // exit action
END_STEP
TRANSITION FROM OpeningDoor TO End
    := SenseOpen;
END_TRANSITION
STEP End:
    _aEnd_active(N);  // step action
    _aEnd_exit(P0);  // exit action
END_STEP
TRANSITION FROM End TO Init
    := NOT Do_;
END_TRANSITION

ACTION _aInit_active:
State := S_Init;
END_ACTION

ACTION _aReady_active:
State := S_Ready;
END_ACTION

ACTION _aBusy_active:
State := S_Busy;
END_ACTION

ACTION _aOpeningDoor_active:
ActOpening := TRUE;
END_ACTION

ACTION _aEnd_active:
Done := TRUE;
END_ACTION

ACTION _aEnd_exit:
Done := FALSE;
END_ACTION

ACTION _aOpeningDoor_exit:
ActOpening := FALSE;
END_ACTION

END_FUNCTION_BLOCK

// Device/Application/GAs/Motor_GA
FUNCTION_BLOCK Motor_GA
VAR_INPUT
	Do_: BOOL;
	DoWhat: DoWhats_Motor;
	SenseRamp: BOOL;
	SenseDeck: BOOL;
	SenseUplimit: BOOL;
	SenseDownlimit: BOOL;
END_VAR
VAR_OUTPUT
	State: State_GA;
	Done: BOOL;
	Fault_State: Fault := None;
	MotorElevator: BOOL;
	Direction: BOOL;
	Velocity: BOOL;
END_VAR
VAR
	Seq_State: SensorSequence := Seq_Deck;
	CheckOk: BOOL;
	FirstDeckPassage : BOOL := TRUE;
END_VAR

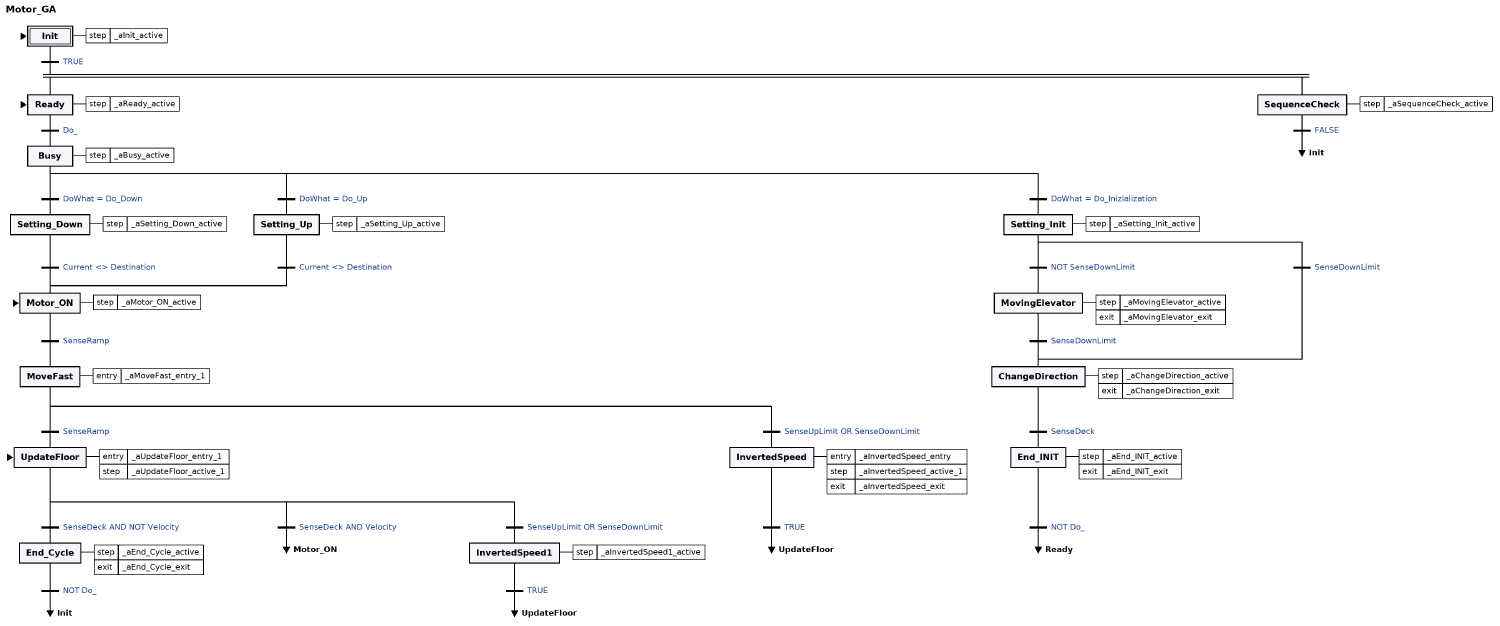
INITIAL_STEP Init:
    _aInit_active(N);  // step action
END_STEP
TRANSITION FROM Init TO (Ready, SequenceCheck)
    := TRUE;
END_TRANSITION
STEP Ready:
    _aReady_active(N);  // step action
END_STEP
STEP SequenceCheck:
    _aSequenceCheck_active(N);  // step action
END_STEP
TRANSITION FROM SequenceCheck TO Init
    := FALSE;
END_TRANSITION
TRANSITION FROM Ready TO Busy
    := Do_;
END_TRANSITION
STEP Busy:
    _aBusy_active(N);  // step action
END_STEP
TRANSITION FROM Busy TO Setting_Down
    := DoWhat = Do_Down;
END_TRANSITION
STEP Setting_Down:
    _aSetting_Down_active(N);  // step action
END_STEP
TRANSITION FROM Setting_Down TO Motor_ON
    := Current <> Destination;
END_TRANSITION
TRANSITION FROM Busy TO Setting_Up
    := DoWhat = Do_Up;
END_TRANSITION
STEP Setting_Up:
    _aSetting_Up_active(N);  // step action
END_STEP
TRANSITION FROM Setting_Up TO Motor_ON
    := Current <> Destination;
END_TRANSITION
TRANSITION FROM Busy TO Setting_Init
    := DoWhat = Do_Inizialization;
END_TRANSITION
STEP Setting_Init:
    _aSetting_Init_active(N);  // step action
END_STEP
TRANSITION FROM Setting_Init TO MovingElevator
    := NOT SenseDownLimit;
END_TRANSITION
STEP MovingElevator:
    _aMovingElevator_active(N);  // step action
    _aMovingElevator_exit(P0);  // exit action
END_STEP
TRANSITION FROM MovingElevator TO ChangeDirection
    := SenseDownLimit;
END_TRANSITION
TRANSITION FROM Setting_Init TO ChangeDirection
    := SenseDownLimit;
END_TRANSITION
STEP ChangeDirection:
    _aChangeDirection_active(N);  // step action
    _aChangeDirection_exit(P0);  // exit action
END_STEP
TRANSITION FROM ChangeDirection TO End_INIT
    := SenseDeck;
END_TRANSITION
STEP End_INIT:
    _aEnd_INIT_active(N);  // step action
    _aEnd_INIT_exit(P0);  // exit action
END_STEP
TRANSITION FROM End_INIT TO Ready
    := NOT Do_;
END_TRANSITION
STEP Motor_ON:
    _aMotor_ON_active(N);  // step action
END_STEP
TRANSITION FROM Motor_ON TO MoveFast
    := SenseRamp;
END_TRANSITION
STEP MoveFast:
    _aMoveFast_entry_1(P1);  // entry action
END_STEP
TRANSITION FROM MoveFast TO UpdateFloor
    := SenseRamp;
END_TRANSITION
TRANSITION FROM MoveFast TO InvertedSpeed
    := SenseUpLimit OR SenseDownLimit;
END_TRANSITION
STEP InvertedSpeed:
    _aInvertedSpeed_entry(P1);  // entry action
    _aInvertedSpeed_active_1(N);  // step action
    _aInvertedSpeed_exit(P0);  // exit action
END_STEP
TRANSITION FROM InvertedSpeed TO UpdateFloor
    := TRUE;
END_TRANSITION
STEP UpdateFloor:
    _aUpdateFloor_entry_1(P1);  // entry action
    _aUpdateFloor_active_1(N);  // step action
END_STEP
TRANSITION FROM UpdateFloor TO End_Cycle
    := SenseDeck AND NOT Velocity;
END_TRANSITION
STEP End_Cycle:
    _aEnd_Cycle_active(N);  // step action
    _aEnd_Cycle_exit(P0);  // exit action
END_STEP
TRANSITION FROM End_Cycle TO Init
    := NOT Do_;
END_TRANSITION
TRANSITION FROM UpdateFloor TO Motor_ON
    := SenseDeck AND Velocity;
END_TRANSITION
TRANSITION FROM UpdateFloor TO InvertedSpeed1
    := SenseUpLimit OR SenseDownLimit;
END_TRANSITION
STEP InvertedSpeed1:
    _aInvertedSpeed1_active(N);  // step action
END_STEP
TRANSITION FROM InvertedSpeed1 TO UpdateFloor
    := TRUE;
END_TRANSITION

ACTION _aBusy_active:
State:= S_Busy;
END_ACTION

ACTION _aEnd_Cycle_active:
MotorElevator := FALSE;
Done := TRUE;
END_ACTION

ACTION _aEnd_INIT_exit:
Done := FALSE;
Seq_State := Seq_Deck;      //dopo Homing, imposto la sequenza dei sensori allo stato iniziale (Seq_Deck)
FirstDeckPassage := FALSE;  //FirstDeckPassege posto a False per evitare che il progetto dia subito errore
END_ACTION

ACTION _aInit_active:
State:= S_Init;
END_ACTION

ACTION _aReady_active:
State:= S_Ready;
END_ACTION

ACTION _aEnd_Cycle_exit:
Done := FALSE;
END_ACTION

ACTION _aMotor_ON_active:
MotorElevator := TRUE;
END_ACTION

ACTION _aSetting_Down_active:
Direction := FALSE;
Velocity  := FALSE;
END_ACTION

ACTION _aMovingElevator_active:
MotorElevator := TRUE;
END_ACTION

ACTION _aSetting_Init_active:
Direction := FALSE;
Velocity  := FALSE;
END_ACTION

ACTION _aSetting_Up_active:
Direction := TRUE;
Velocity  := FALSE;
END_ACTION

ACTION _aUpdateFloor_active_1:
IF (Current = Destination) THEN
	Velocity := FALSE;
END_IF
END_ACTION

ACTION _aEnd_INIT_active:
Done := TRUE;
END_ACTION

ACTION _aChangeDirection_exit:
MotorElevator := FALSE;
Current := 0;  // finito Homing, imposto piano corrente a 0, 
			   //in modo tale da sapere il piano da cui parto per eventuali nuove chiamate successive.
END_ACTION

ACTION _aChangeDirection_active:
MotorElevator := TRUE;
Direction := TRUE;
END_ACTION

ACTION _aMovingElevator_exit:
MotorElevator := FALSE;
END_ACTION

ACTION _aSequenceCheck_active:
// Gestione passaggio della cabina attraverso le rampe e i piani. Utilizzo Seq_State per verificare la sequenza: Deck → Ramp1 → Ramp2 → Deck.
// In caso di incongruenze tra i sensori e lo stato atteso, viene rilevato un guasto e il sistema entra nello stato Seq_Fault.
// La variabile CheckOk serve per abilitare l’avanzamento nella sequenza e viene resettata dopo ogni transizione.

IF CheckOk THEN
	IF Seq_State = Seq_Deck THEN
		IF SenseRamp THEN
			Seq_State := Seq_Ramp1;
			CheckOk := FALSE;
	    ELSIF SenseDeck AND Motor_GA_0.DoWhat <> Do_Inizialization AND FirstDeckPassage THEN        //FirstDeckPassage permette di tollerare il primo rilevamento 
			Fault_State := MagnetRamp;																//del sensore di piano (SenseDeck) subito dopo l’inizializzazione. 																					
			CheckOk := FALSE;																		//Dopo questo evento, rilevamenti incoerenti verranno considerati come fault.
		END_IF																						
		
	ELSIF Seq_State = Seq_Ramp1 THEN             
		IF SenseRamp THEN
			Seq_State := Seq_Ramp2;
			CheckOk := FALSE;
		ELSIF SenseDeck AND Motor_GA_0.DoWhat <> Do_Inizialization  THEN
			Seq_State := Seq_Fault;
			Fault_State := MagnetRamp;
			IF Motor_GA_0.DoWhat = Do_Up THEN
				Current := Current + 1;
			ELSIF Motor_GA_0.DoWhat = Do_Down THEN
				Current := Current - 1;
			END_IF
			CheckOk := FALSE;
		END_IF
	
	ELSIF Seq_State = Seq_Ramp2 THEN             
		IF SenseDeck THEN
			Seq_State := Seq_Deck;
			CheckOk := FALSE;
		ELSIF (SenseRamp OR SenseUpLimit OR SenseDownLimit) AND Motor_GA_0.DoWhat <> Do_Inizialization THEN          //OR SenseUpLimit OR SenseDownLimit
			Seq_State := Seq_Fault;
			Fault_State := MagnetDeck;
			IF Motor_GA_0.DoWhat = Do_Up THEN
				Current := Current + 1;
			ELSIF Motor_GA_0.DoWhat = Do_Down THEN
				Current := Current - 1;
			END_IF
			CheckOk := FALSE;
		END_IF
	END_IF
END_IF

IF NOT SenseDeck AND NOT SenseRamp AND Fault_State = None THEN
	CheckOk := TRUE;
END_IF
END_ACTION

ACTION _aMoveFast_entry_1:
Velocity := TRUE;
END_ACTION

ACTION _aUpdateFloor_entry_1:
// Aggiornamento del piano corrente in base alla direzione di marcia. 
// Aggiornamento avviene nel sensore di rampa che antecede il sensore del piano successivo.
IF(NOT Direction) THEN
	Current := Current - 1;
ELSE
	Current := Current + 1;
END_IF
END_ACTION

ACTION _aInvertedSpeed1_active:
// Inversione della direzione in caso di Fault Deck ai piani estremi (0 o 7)

IF Motor_GA_0.DoWhat = Do_Down THEN
	Direction := TRUE;
	ELSIF Motor_GA_0.DoWhat = Do_Up THEN
		Direction := FALSE;
END_IF
END_ACTION

ACTION _aInvertedSpeed_active_1:
// Caso particolare per i piani G e 7 nel caso di RampFault
IF Motor_GA_0.DoWhat = Do_Down THEN
	Direction := TRUE;
	ELSIF Motor_GA_0.DoWhat = Do_Up THEN
		Direction := FALSE;
END_IF
END_ACTION

ACTION _aInvertedSpeed_exit:
// Correzione dell'aggiornamento del Current nel caso di inversione della direzione causata da fault (MagnetRamp) ai piani estremi (0 o 7). 
// La logica di SequenceCheck ha aggiornato Current nella direzione sbagliata (quella precedente). 
// Questo blocco annulla e corregge l’errore, riportando Current al valore corretto.

IF(NOT Direction) THEN
	Current := Current + 1;
ELSE
	Current := Current - 1;
END_IF
END_ACTION

ACTION _aInvertedSpeed_entry:
IF(NOT Direction) THEN
	Current := Current - 1;
ELSE
	Current := Current + 1;
END_IF
END_ACTION

END_FUNCTION_BLOCK

// Device/Application/Visualization
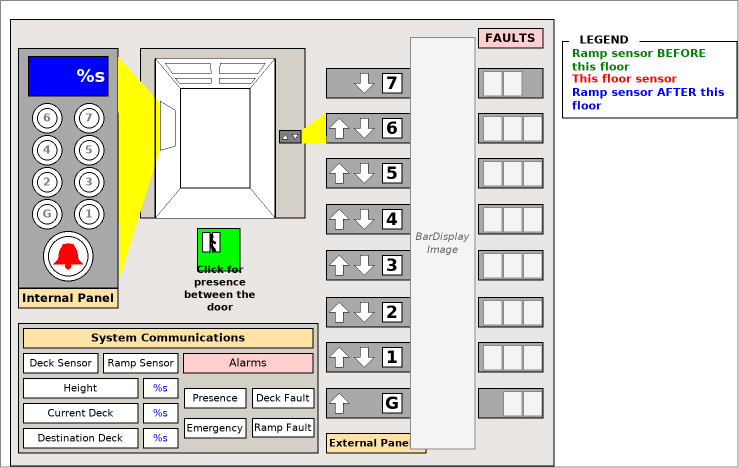
VISUALIZATION Visualization  // 739x468
    Rectangle (10,19 544x447)
    Rectangle (197,228 43x43), colour toggle: GVL.Presence
    Rectangle (18,323 300x130)
    Rectangle (326,433 100x20), "External Panels"
    Rectangle (326,342 100x30)
    Rectangle (382,347 20x20), "1"
    Polygon (354,357) (360,357) (360,347) (368,347) (368,357) (374,357) (364,367), colour toggle: GVL.DownDeck1Vis
        tap GVL.DownDeck1
    Polygon (329,357) (335,357) (335,367) (343,367) (343,357) (349,357) (339,347), colour toggle: GVL.UpDeck1Vis
        tap GVL.UpDeck1
    Rectangle (326,297 100x30)
    Rectangle (382,302 20x20), "2"
    Polygon (354,312) (360,312) (360,302) (368,302) (368,312) (374,312) (364,322), colour toggle: GVL.DownDeck2Vis
        tap GVL.DownDeck2
    Polygon (329,312) (335,312) (335,322) (343,322) (343,312) (349,312) (339,302), colour toggle: GVL.UpDeck2Vis
        tap GVL.UpDeck2
    Rectangle (326,250 100x30)
    Rectangle (382,255 20x20), "3"
    Polygon (354,265) (360,265) (360,255) (368,255) (368,265) (374,265) (364,275), colour toggle: GVL.DownDeck3Vis
        tap GVL.DownDeck3
    Polygon (329,265) (335,265) (335,275) (343,275) (343,265) (349,265) (339,255), colour toggle: GVL.UpDeck3Vis
        tap GVL.UpDeck3
    Rectangle (326,204 100x30)
    Rectangle (382,209 20x20), "4"
    Polygon (354,219) (360,219) (360,209) (368,209) (368,219) (374,219) (364,229), colour toggle: GVL.DownDeck4Vis
        tap GVL.DownDeck4
    Polygon (329,219) (335,219) (335,229) (343,229) (343,219) (349,219) (339,209), colour toggle: GVL.UpDeck4Vis
        tap GVL.UpDeck4
    Rectangle (326,158 100x30)
    Rectangle (382,163 20x20), "5"
    Polygon (354,173) (360,173) (360,163) (368,163) (368,173) (374,173) (364,183), colour toggle: GVL.DownDeck5Vis
        tap GVL.DownDeck5
    Polygon (329,173) (335,173) (335,183) (343,183) (343,173) (349,173) (339,163), colour toggle: GVL.UpDeck5Vis
        tap GVL.UpDeck5
    Rectangle (326,113 100x30)
    Rectangle (382,118 20x20), "6"
    Polygon (354,128) (360,128) (360,118) (368,118) (368,128) (374,128) (364,138), colour toggle: GVL.DownDeck6Vis
        tap GVL.DownDeck6
    Polygon (329,128) (335,128) (335,138) (343,138) (343,128) (349,128) (339,118), colour toggle: GVL.UpDeck6Vis
        tap GVL.UpDeck6
    Rectangle (326,68 100x30)
    Rectangle (382,73 20x20), "7"
    Polygon (354,83) (360,83) (360,73) (368,73) (368,83) (374,83) (364,93), colour toggle: GVL.DownDeck7Vis
        tap GVL.DownDeck7
    Rectangle (326,388 100x30)
    Rectangle (382,393 20x20), "G"
    Polygon (329,403) (335,403) (335,413) (343,413) (343,403) (349,403) (339,393), colour toggle: GVL.UpDeckGVis
        tap GVL.UpDeckG
    RoundedRectangle (18,48 100x240)
    Rectangle (18,288 100x20), "Internal Panel"
    Ellipse (74,199 30x30), colour toggle: GVL.P1Vis
    Ellipse (79,204 20x20), "1"
        tap GVL.P1
    Ellipse (32,199 30x30), colour toggle: GVL.PGVis
    Ellipse (37,204 20x20), "G"
        tap GVL.PG
    Ellipse (74,167 30x30), colour toggle: GVL.P3Vis
    Ellipse (79,172 20x20), "3"
        tap GVL.P3
    Ellipse (32,167 30x30), colour toggle: GVL.P2Vis
    Ellipse (37,172 20x20), "2"
        tap GVL.P2
    Ellipse (74,135 30x30), colour toggle: GVL.P5Vis
    Ellipse (79,140 20x20), "5"
        tap GVL.P5
    Ellipse (32,135 30x30), colour toggle: GVL.P4Vis
    Ellipse (37,140 20x20), "4"
        tap GVL.P4
    Ellipse (74,103 30x30), colour toggle: GVL.P7Vis
    Ellipse (79,108 20x20), "7"
        tap GVL.P7
    Ellipse (32,103 30x30), colour toggle: GVL.P6Vis
    Ellipse (37,108 20x20), "6"
        tap GVL.P6
    Rectangle (28,56 80x40), "%s", text variable: GVL.Destination
    Ellipse (43,231 50x50), tooltip "EMERGENCY", colour toggle: GVL.Emergency
    Group (48,236 40x40)
        toggle GVL.Emergency
        Ellipse (0,0 40x40), tooltip "EMERGENCY"
        Polygon (5,28) (10,23) (11,15) (15,8) (20,7) (25,8) (29,15) (30,23) (35,28)
        Ellipse (17,27 6x6)
    Polygon (35,72) (45,62) (55,72), colour toggle: GVL.Motor_on AND GVL.Up
    Polygon (35,80) (45,90) (55,80), colour toggle: GVL.Motor_on AND NOT GVL.Up
    Group (140,48 165x170)
        Rectangle (0,0 165x170)
        Rectangle (15,10 120x160)
        Polygon (40,40) (15,10) (135,10) (110,40)
        Rectangle (40,40 70x100)
        Polygon (15,170) (40,140) (110,140) (135,170)
        Polygon (20,102) (20,53) (35,62) (35,98)
        Polygon (79,35) (79,30) (115,30) (111,35)
        Polygon (39,35) (35,30) (71,30) (71,35)
        Polygon (32,25) (25,15) (70,15) (71,25)
        Polygon (79,25) (80,15) (125,15) (118,25)
        Group (139,82 22x13)
            Rectangle (0,0 22x13)
            Polygon (3,9) (6,4) (9,9)
            Polygon (13,4) (16,9) (19,4)
    BarDisplayImage (410,37 65x412), value: GVL.Height, style: BarDisplayImage-Gray, scale format: %.0f, scale -20..160
        p3451962224: VisuNativeControl.IP_Offline.Browser
    Rectangle (478,68 65x30)
    Rectangle (478,342 65x30)
    Rectangle (478,297 65x30)
    Rectangle (478,250 65x30)
    Rectangle (478,204 65x30)
    Rectangle (478,158 65x30)
    Rectangle (478,113 65x30)
    Rectangle (478,388 65x30)
    RockerSwitch (483,345 19x25), variable: GVL.Ramp1Down, behaviour: TOGGLE, style: Switch-RockerSwitch-Green
    RockerSwitch (503,345 19x25), variable: GVL.Sensor1, behaviour: TOGGLE, style: Switch-RockerSwitch-Red
    RockerSwitch (523,345 19x25), variable: GVL.Ramp1Up, behaviour: TOGGLE, style: Switch-RockerSwitch-Blue
    RockerSwitch (483,300 19x25), variable: GVL.Ramp2Down, behaviour: TOGGLE, style: Switch-RockerSwitch-Green
    RockerSwitch (503,300 19x25), variable: GVL.Sensor2, behaviour: TOGGLE, style: Switch-RockerSwitch-Red
    RockerSwitch (523,300 19x25), variable: GVL.Ramp2Up, behaviour: TOGGLE, style: Switch-RockerSwitch-Blue
    RockerSwitch (483,253 19x25), variable: GVL.Ramp3Down, behaviour: TOGGLE, style: Switch-RockerSwitch-Green
    RockerSwitch (503,253 19x25), variable: GVL.Sensor3, behaviour: TOGGLE, style: Switch-RockerSwitch-Red
    RockerSwitch (523,253 19x25), variable: GVL.Ramp3Up, behaviour: TOGGLE, style: Switch-RockerSwitch-Blue
    RockerSwitch (483,207 19x25), variable: GVL.Ramp4Down, behaviour: TOGGLE, style: Switch-RockerSwitch-Green
    RockerSwitch (503,207 19x25), variable: GVL.Sensor4, behaviour: TOGGLE, style: Switch-RockerSwitch-Red
    RockerSwitch (523,207 19x25), variable: GVL.Ramp4Up, behaviour: TOGGLE, style: Switch-RockerSwitch-Blue
    RockerSwitch (483,161 19x25), variable: GVL.Ramp5Down, behaviour: TOGGLE, style: Switch-RockerSwitch-Green
    RockerSwitch (503,161 19x25), variable: GVL.Sensor5, behaviour: TOGGLE, style: Switch-RockerSwitch-Red
    RockerSwitch (523,161 19x25), variable: GVL.Ramp5Up, behaviour: TOGGLE, style: Switch-RockerSwitch-Blue
    RockerSwitch (483,116 19x25), variable: GVL.Ramp6Down, behaviour: TOGGLE, style: Switch-RockerSwitch-Green
    RockerSwitch (503,116 19x25), variable: GVL.Sensor6, behaviour: TOGGLE, style: Switch-RockerSwitch-Red
    RockerSwitch (523,116 19x25), variable: GVL.Ramp6Up, behaviour: TOGGLE, style: Switch-RockerSwitch-Blue
    RockerSwitch (483,71 19x25), variable: GVL.Ramp7Down, behaviour: TOGGLE, style: Switch-RockerSwitch-Green
    RockerSwitch (503,71 19x25), variable: GVL.Sensor7, behaviour: TOGGLE, style: Switch-RockerSwitch-Red
    RockerSwitch (503,391 19x25), variable: GVL.SensorG, behaviour: TOGGLE, style: Switch-RockerSwitch-Red
    RockerSwitch (523,391 19x25), variable: GVL.RampGUp, behaviour: TOGGLE, style: Switch-RockerSwitch-Blue
    Rectangle (478,28 65x20), "FAULTS"
    Polygon (302,130) (325,113) (326,143) (302,143), invisible if: (GVL.Closing OR GVL.Opening) OR GVL.Closed
    Polygon (118,57) (159,102) (159,151) (119,279), invisible if: (GVL.Closing OR GVL.Opening) OR GVL.Closed
    Rectangle (155,58 0x160)
        p3528305787: GVL.Door
    Rectangle (275,58 0x160)
        p3528305787: -GVL.Door
    Rectangle (23,328 290x20), "System Communications"
    Rectangle (183,353 130x20), "Alarms"
    Rectangle (23,353 75x20), "Deck Sensor", colour toggle: GVL.DeckSensor
    Rectangle (143,378 35x20), "%s", text variable: GVL.Height
    Rectangle (184,388 62x20), "Presence", colour toggle: GVL.Presence
    Rectangle (103,353 75x20), "Ramp Sensor", colour toggle: GVL.RampSensor
    Rectangle (143,403 35x20), "%s", text variable: GVL.Current
    Rectangle (143,428 35x20), "%s", text variable: GVL.Destination
    Rectangle (252,388 62x20), "Deck Fault", colour toggle: GVL.FaultSensorAlarm
    Rectangle (184,418 62x20), "Emergency", colour toggle: GVL.EmergencyVis
    Rectangle (252,418 62x19), "Ramp Fault", colour toggle: GVL.FaultRampAlarm
    Rectangle (23,378 115x20), "Height"
    Rectangle (23,403 115x20), "Current Deck"
    Rectangle (23,428 115x20), "Destination Deck"
    Group (562,25 175x93)
        Rectangle (0,16 175x77)
        Rectangle (7,39 160x30), "This floor sensor"
        Rectangle (7,59 160x30), "Ramp sensor AFTER this floor"
        Rectangle (7,0 70x30), "LEGEND"
        Rectangle (7,20 160x30), "Ramp sensor BEFORE this floor"
    Group (202,232 33x34)
        toggle GVL.Presence
        Rectangle (10,0 8x20)
        Polygon (5,10) (12,20) (14,18) (5,6)
        Ellipse (6,2 5x5)
        Polygon (4,8) (13,12) (14,10) (4,4)
        Rectangle (0,0 8x20)
    Rectangle (169,273 102x31), "Click for presence between the door"
END_VISUALIZATION
